TYPE ST_EL3214CoeReadData :
STRUCT
	wIdx: WORD;
	bySubIdx: BYTE;
	bReadOK: BOOL;
	dwData: DWORD;
	nSize: UDINT;
END_STRUCT
END_TYPE

(* stored: Version 1.1.0.1, ProductVersion 3.1.4024.15
   DUT ST_EL3214CoeReadData: Id {d774c257-9d55-485e-bfa8-c857cde7352d} *)
